Fanuc KAREL source: ko00075.KL

-- PROVISIONAL review KL for V770-1; original PC SHA256 be8bdcc7a4e7251bf4c39d9a619dd2ead7e7a2d9249e57a2a622d04e6750e107
-- Incomplete behavior may be omitted. Consult companion uncertainty JSON. Do not deploy.
PROGRAM KO00075
%NOLOCKGROUP
BEGIN
  -- UNRESOLVED_PC offsets 5-12; opcodes 9D,23
  -- UNRESOLVED_PC offsets 17-66; opcodes 27,22,1C,27,49,7E,AD,22,31,7E,4A
  -- UNRESOLVED_PC offsets 71-75; opcodes 7F
END KO00075
